FUNCTION_BLOCK Controle_PID (* Parametros de PID (padrao PID do legado); o pidCtl fica no processo *)
  (* Standard: 61499-2 *)
  (* Version 1.0, 21/10/2026, Hidryco, Hidryco, 1.0: Parametros de PID (padrao PID do legado); o pidCtl fica no processo *)
  PACKAGE Hidryco.HidrycoLib;
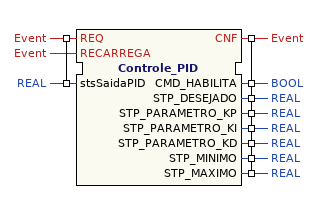
  EVENT_INPUT
    REQ WITH stsSaidaPID; (* Status vindo do processo *)
    RECARREGA; (* Reenvia os ajustes persistentes (chamado no fim do INIT do processo) *)
  END_EVENT
  EVENT_OUTPUT
    CNF WITH CMD_HABILITA, STP_DESEJADO, STP_PARAMETRO_KP, STP_PARAMETRO_KI, STP_PARAMETRO_KD, STP_MINIMO, STP_MAXIMO; (* Ajustes para o processo (mudanca na IHM, OPC UA ou recarga) *)
  END_EVENT
  VAR_INPUT
    stsSaidaPID : REAL; (* Saida do PID (%) *)
  END_VAR
  VAR_OUTPUT
    CMD_HABILITA : BOOL; (* PID habilitado *)
    STP_DESEJADO : REAL; (* Valor desejado *)
    STP_PARAMETRO_KP : REAL; (* Ganho (Kp) *)
    STP_PARAMETRO_KI : REAL; (* Tempo integral (s) *)
    STP_PARAMETRO_KD : REAL; (* Tempo derivativo (s) *)
    STP_MINIMO : REAL; (* Saída mínima *)
    STP_MAXIMO : REAL; (* Saída máxima *)
  END_VAR
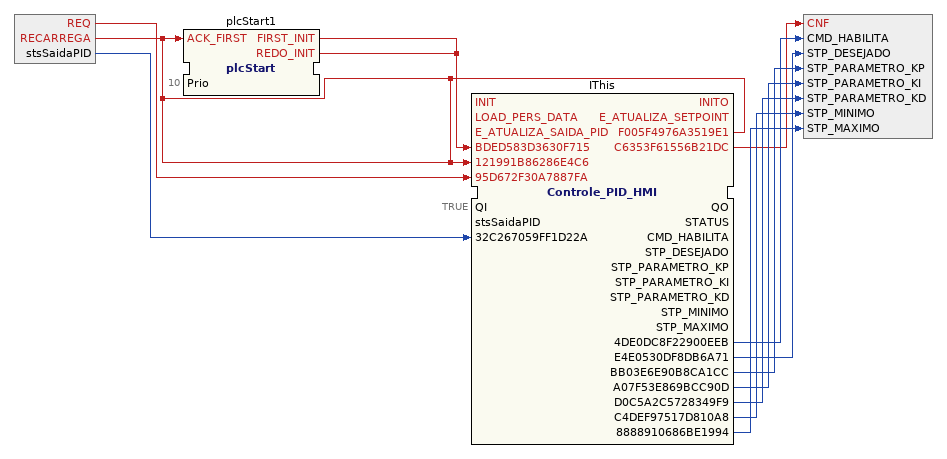
  FBS
    IThis : Controle_PID_HMI(QI := TRUE);
    plcStart1 : plcStart(Prio := 10);
  END_FBS
  EVENT_CONNECTIONS
    plcStart1.FIRST_INIT TO IThis.BDED583D3630F715;
    plcStart1.REDO_INIT TO IThis.BDED583D3630F715;
    IThis.F005F4976A3519E1 TO IThis.121991B86286E4C6;
    IThis.F005F4976A3519E1 TO plcStart1.ACK_FIRST;
    RECARREGA TO IThis.121991B86286E4C6;
    IThis.C6353F61556B21DC TO CNF;
    REQ TO IThis.95D672F30A7887FA;
  END_CONNECTIONS
  DATA_CONNECTIONS
    IThis.4DE0DC8F22900EEB TO CMD_HABILITA;
    IThis.E4E0530DF8DB6A71 TO STP_DESEJADO;
    IThis.BB03E6E90B8CA1CC TO STP_PARAMETRO_KP;
    IThis.A07F53E869BCC90D TO STP_PARAMETRO_KI;
    IThis.D0C5A2C5728349F9 TO STP_PARAMETRO_KD;
    IThis.C4DEF97517D810A8 TO STP_MINIMO;
    IThis.8888910686BE1994 TO STP_MAXIMO;
    stsSaidaPID TO IThis.32C267059FF1D22A;
  END_CONNECTIONS
END_FUNCTION_BLOCK
